TYPE ST_ConfigConveyor :
STRUCT
	(* vo_Config of _FB_ConfigConveyor: the gateway writes stStaging and stStaged, reads stStatus and stActive. *)
	stStaging : ST_ConfigStaging;
	stStaged : ST_ConfigConveyorParam;
	stStatus : ST_ConfigStatus;
	stActive : ST_ConfigConveyorParam; // effective values: the active set while one is valid, else the program values
END_STRUCT
END_TYPE

(* stored: Version 1.1.0.1
   DUT ST_ConfigConveyor: Id {6b07eba1-2622-4d46-b88d-ba87be036220} *)
